// TIA Portal V21 export
FUNCTION_BLOCK "FbdLogic"   // FB13, FBD
TITLE = Function block logic
{ S7_Optimized_Access := 'TRUE' }
// Bit logic in function block diagram: gates, a set and reset box, an edge and a jump.
   VAR_INPUT
      start : Bool;
      stop : Bool;
      door : Bool;
   END_VAR
   VAR_OUTPUT
      motor : Bool;
      lamp : Bool;
      fault : Bool;
   END_VAR
   VAR
      latched : Bool;
      edgeMemory : Bool;
   END_VAR
   VAR_TEMP   // added for the SCL form of the ladder/FBD networks
      _w1 : Bool;
   END_VAR
BEGIN

REGION Network 1: Start and stop
   // OR and AND boxes drive the motor, stop negated.
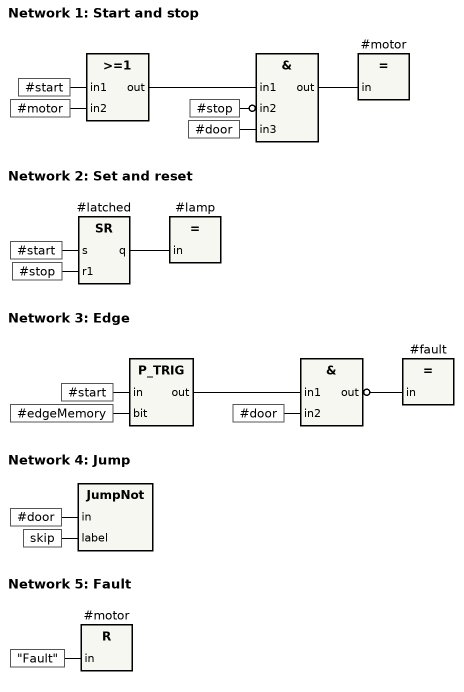
   #motor := (#start OR #motor) AND NOT #stop AND #door;
END_REGION

REGION Network 2: Set and reset
   // A set and reset box, its output on the lamp.
   IF #start THEN
       #latched := TRUE;   // SR flip-flop
   END_IF;
   IF #stop THEN #latched := FALSE; END_IF;
   #lamp := #latched;
END_REGION

REGION Network 3: Edge
   // A rising edge of start and the door, negated, is the fault.
   #_w1 := #start AND NOT #edgeMemory;   // rising edge
   #edgeMemory := #start;
   #fault := NOT (#_w1 AND #door);
END_REGION

REGION Network 4: Jump
   // Without the door closed, skip to the end.
   // no SCL statement known for JumpNot: written as a call
   JumpNot(in := #door, label := skip);
END_REGION

REGION Network 5: Fault
   // Jump target; a fault resets the motor.
   skip:
   IF "Fault" THEN #motor := FALSE; END_IF;
END_REGION
END_FUNCTION_BLOCK
